// TIA Portal V21 export
TYPE "UDT_Recipe"
TITLE = Filling recipe
   STRUCT
      Id : Int := 1;   // Recipe number
      RecipeName : String[20] := 'Default';   // Recipe name
      Volumes : Array[1..10] of Real;   // Volume per filling step in litres
      FillTime : Time := T#5S;   // Maximum filling time per step
      Temperature : Real := 20.0;   // Product temperature in degrees Celsius
   END_STRUCT;
   // Volumes[1] := 1.0;
   // Volumes[2] := 2.0;
   // Volumes[3..10] := 0.5;
END_TYPE
